// TIA Portal V20 export
FUNCTION_BLOCK "Ampelbaustein_MG"   // FB145, STL
{ S7_Optimized_Access := 'FALSE' }
// stored: AutoNumber false
   VAR_INPUT
      Sammelstoerung : Bool;
      BA_0 : Bool;
      BA_A : Bool;
      BA_M : Bool;
      BA_R : Bool;
      BA_V : Bool;
      Ablauf_ist_aktiv : Bool;
      Blinker : Bool;
   END_VAR
   VAR_OUTPUT
      Ampel_rot : Bool;
      Ampel_gelb : Bool;
      Ampel_gruen : Bool;
      Akkustik : Bool;
   END_VAR
   VAR
      Timer_Hupe_EIN { S7_SetPoint := 'True'} : TON_TIME;
      Timer_Hupe_Aus { S7_SetPoint := 'True'} : TON_TIME;
      Ampel_Zustand : Int;
   END_VAR
BEGIN

NETWORK
TITLE = Ampel Betriebsart 0-4
      L     0;
      T     #Ampel_Zustand;

// Grün
      A     #Ablauf_ist_aktiv;
      A     #BA_A;
      AN    #Sammelstoerung;
      JCN   zustand_rot;
      L     1;
      T     #Ampel_Zustand;
      JU    auswertung;

// Rot
zustand_rot:NOP   0;
      A     #Sammelstoerung;
      JCN   zustand_gelb;
      L     2;
      T     #Ampel_Zustand;
      JU    auswertung;


// Gelb
zustand_gelb:NOP   0;
      A     #BA_A;
      O     #BA_M;
      O     #BA_V;
      O     #BA_R;
      JCN   auswertung;
      L     3;
      T     #Ampel_Zustand;

// Aus
zustand_Aus:NOP   0;
      A     #BA_0;
      JCN   auswertung;
      L     4;
      T     #Ampel_Zustand;





NETWORK
TITLE = Sprungliste in die jewilige Ampelbeschaltung (wie case anweisung)
auswertung:NOP   0;
      L     #Ampel_Zustand;
      JL    end;
      JU    NOP;
      JU    grün;
      JU    rot;
      JU    gelb;
      JU    Aus;
end:  JU    ENDE;

NETWORK
TITLE = Nicht definiert
NOP:  NOP   0;


      CLR;
      =     #Ampel_gelb;
      =     #Ampel_rot;
      =     #Ampel_gruen;
      =     #Akkustik;



      JU    ENDE;


NETWORK
TITLE = Grün
grün: NOP   0;
      SET;
      =     #Ampel_gruen;
      CLR;
      =     #Ampel_gelb;
      =     #Ampel_rot;
      =     #Akkustik;
      JU    ENDE;


NETWORK
TITLE = Rot
rot:  NOP   0;
      SET;
      =     #Ampel_rot;
      CLR;
      =     #Ampel_gelb;
      =     #Ampel_gruen;
      =     #Akkustik;
      JU    ENDE;

NETWORK
TITLE = Gelb
gelb: NOP   0;
      SET;
      =     #Ampel_gelb;
      CLR;
      =     #Ampel_rot;
      =     #Ampel_gruen;
      =     #Akkustik;

      JU    ENDE;

NETWORK
TITLE = Aus
Aus:  NOP   0;
      SET;

      CLR;
      =     #Ampel_rot;
      =     #Ampel_gelb;
      =     #Ampel_gruen;
      =     #Akkustik;

      JU    ENDE;

NETWORK
TITLE = ENDE Sprungleiste
ENDE: NOP   0;


NETWORK
TITLE = Störungshupe
      CALL  #Timer_Hupe_EIN
      ( IN := #Sammelstoerung,
        PT := T#5M,
        Q  := ,
        ET := 
      );

      CALL  #Timer_Hupe_Aus
      ( IN := #Sammelstoerung,
        PT := T#10M,
        Q  := ,
        ET := 
      );

      A     #Sammelstoerung;
      A     #Blinker;
//      U     #Timer_Hupe_EIN.Q
//      UN    #Timer_Hupe_Aus.Q
      A     #BA_A;
      =     #Akkustik;

END_FUNCTION_BLOCK
